FUNCTION_BLOCK DiagSetDTC (* Activate or deactivate a diagnostic trouble code (DTC) in the DM1 message *)
  (* Standard: 61499-2; Description: Calls iso_BaseDiagSetDM1DTC() of the CCI ISOBUS driver (ISO 11783-12). \n The driver sends DM1 once per second while a DTC is active, keeps the occurrence count \n and handles DM2 (previously active DTCs) and DM3 (clear) by itself. \n Every activation of an inactive DTC increases the occurrence count. \n s16CfHandle is the handle of an own (internal) CF, e.g. sNetEv.s16Handle of NmGetCfInfo with member thisMember. \n Requires ISO_DIAG_ENABLE_DM1 in the firmware, otherwise s16Status is E_CONFIG. *)
  (* Version 1.0, 2026-11-17, Franz Höpfinger, initial API and implementation and/or initial documentation *)
  PACKAGE isobus::pgn::diag;
  IMPORT isobus::pgn::HANDLE::UNVALID;
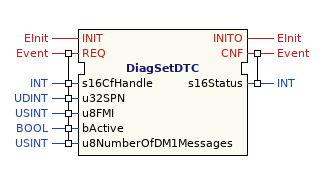
  EVENT_INPUT
    INIT : EInit; (* Service Initialization *)
    REQ WITH s16CfHandle, u32SPN, u8FMI, bActive, u8NumberOfDM1Messages; (* Set the DTC (activate or deactivate) *)
  END_EVENT
  EVENT_OUTPUT
    INITO : EInit; (* Initialization Confirm *)
    CNF WITH s16Status; (* Confirmation *)
  END_EVENT
  VAR_INPUT
    s16CfHandle : INT := UNVALID; (* Handle of the own (internal) CF *)
    u32SPN : UDINT; (* Suspect Parameter Number of the trouble code (19 bit) *)
    u8FMI : USINT; (* Failure Mode Identifier, see isobus::pgn::diag::FMI *)
    bActive : BOOL; (* TRUE = activate, FALSE = deactivate the DTC *)
    u8NumberOfDM1Messages : USINT; (* 0 or 255: active until deactivated; 1..254: deactivate automatically after this number of DM1 messages (seconds) *)
  END_VAR
  VAR_OUTPUT
    s16Status : INT; (* Return value of iso_BaseDiagSetDM1DTC(): 0 = OK, < 0 = error *)
  END_VAR
END_FUNCTION_BLOCK
